PROGRAM Counters
  VAR
    h01_a : BOOL;
    CTU0 : CTU;
    h01_q : BOOL;
    h01_b : BOOL;
    h01_c : BOOL;
    h01_d : BOOL;
    h01_cv : INT;
    h02_a : BOOL;
    CTUD0 : CTUD;
    h02_qu : BOOL;
    h02_b : BOOL;
    h02_c : BOOL;
    h02_d : BOOL;
    h02_e : BOOL;
    h02_g : BOOL;
    h02_f : BOOL;
    h02_h : BOOL;
    h02_i : BOOL;
    h02_k : BOOL;
    h02_j : BOOL;
    h02_qd : BOOL;
    h02_cv : INT;
    h03_a : BOOL;
    SR0 : SR;
    h03_q1 : BOOL;
    h03_c : BOOL;
    h03_b : BOOL;
    h03_d : BOOL;
    h03_e : BOOL;
    RS0 : RS;
    h03_q2 : BOOL;
    h03_f : BOOL;
    h03_h : BOOL;
    h03_g : BOOL;
    h04_e : BOOL;
    TON0 : TON;
    h04_q : BOOL;
    h04_a : BOOL;
    h04_b : BOOL;
    h04_c : BOOL;
    h04_d : BOOL;
    h04_et : TIME;
  END_VAR

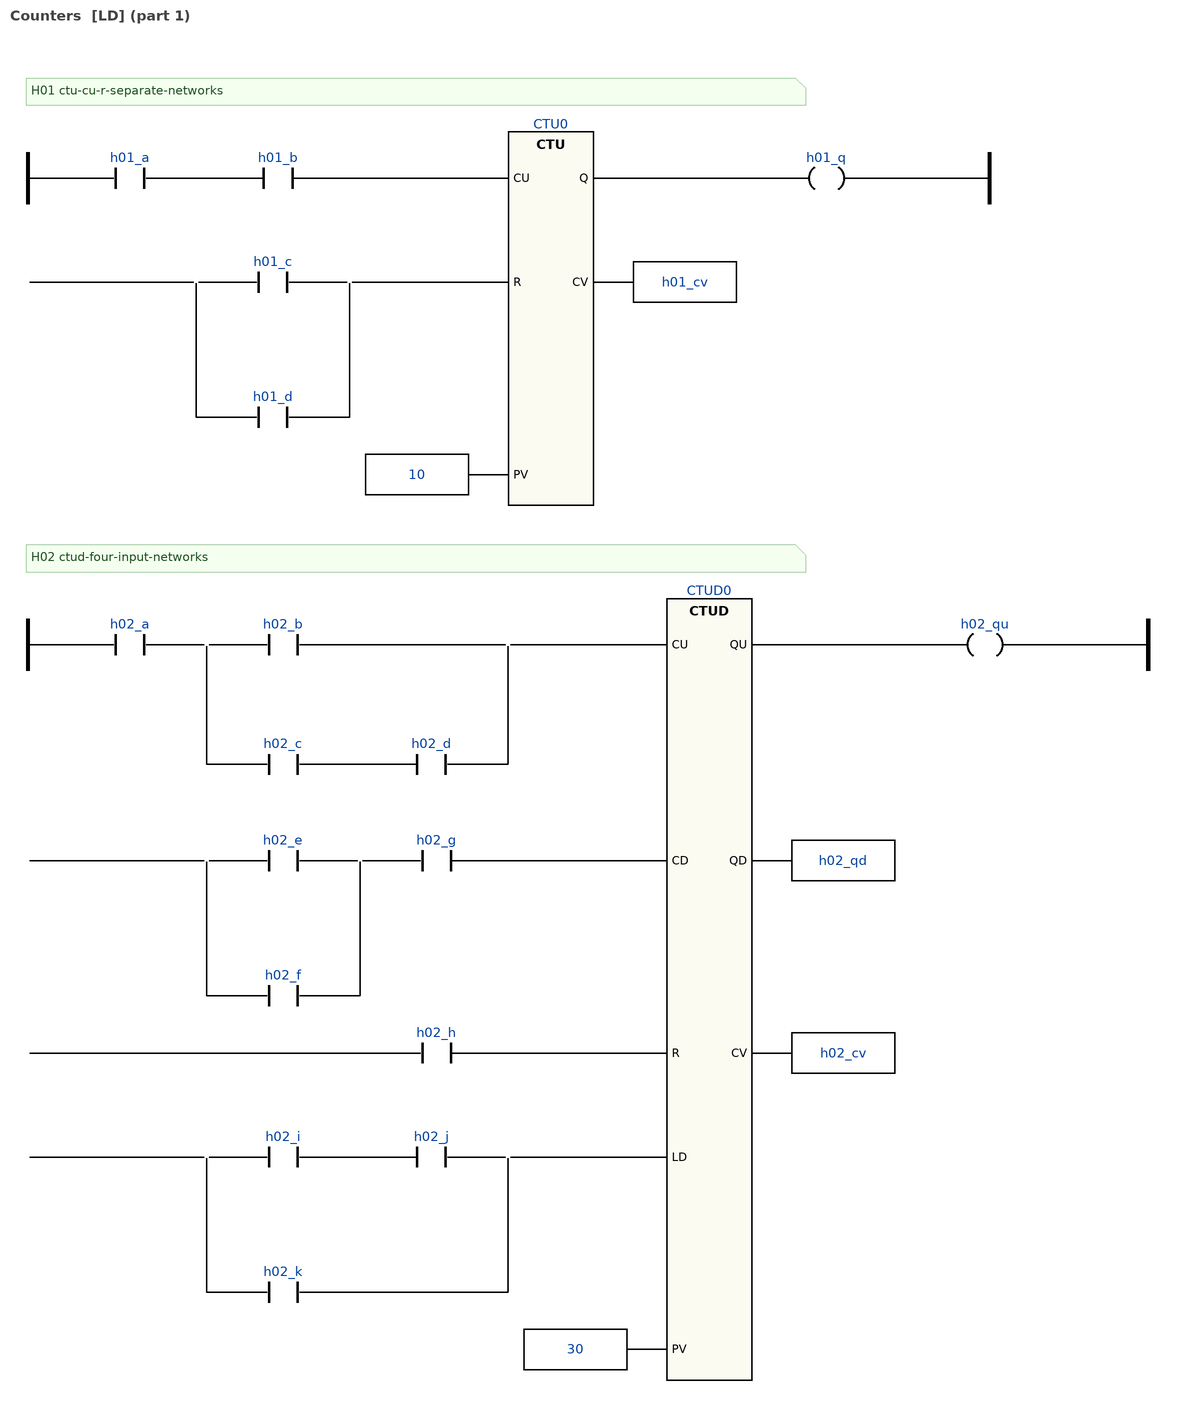
(* LD diagram, written out as Structured Text *)
(* H01 ctu-cu-r-separate-networks *)
CTU0(CU := h01_a AND h01_b, R := h01_c OR h01_d, PV := 10);
h01_q := CTU0.Q;
h01_cv := CTU0.CV;
(* H02 ctud-four-input-networks *)
CTUD0(CU := h02_a AND (h02_b OR h02_c AND h02_d), CD := (h02_e OR h02_f) AND h02_g, R := h02_h, LD := h02_k OR h02_i AND h02_j, PV := 30);
h02_qu := CTUD0.QU;
h02_qd := CTUD0.QD;
h02_cv := CTUD0.CV;
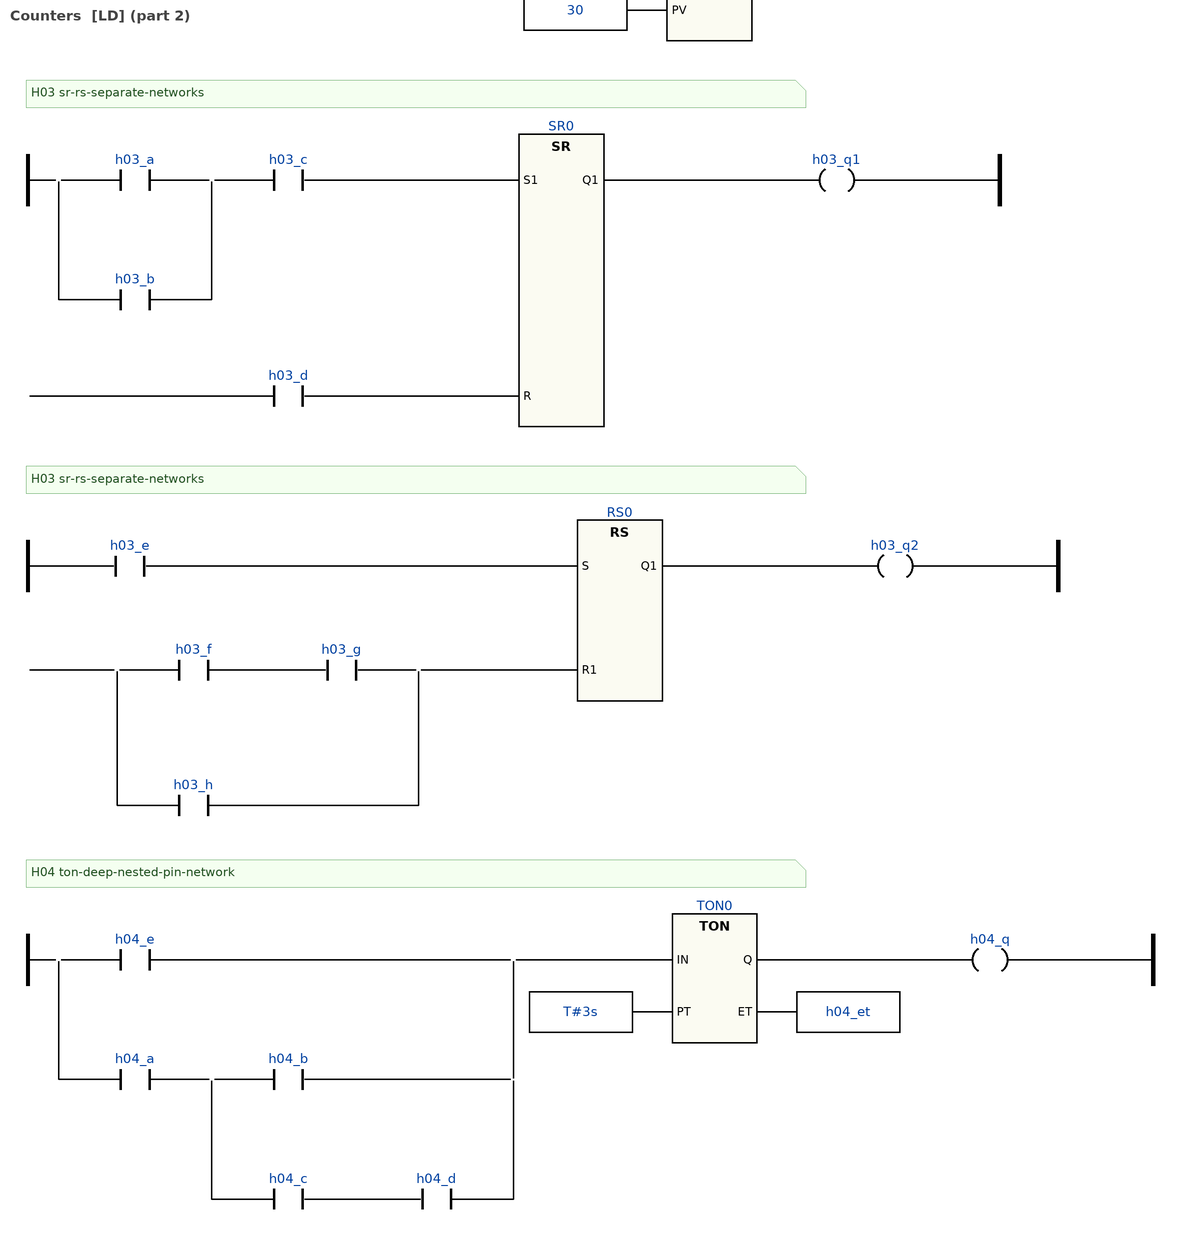
(* H03 sr-rs-separate-networks *)
SR0(S1 := (h03_a OR h03_b) AND h03_c, R := h03_d);
h03_q1 := SR0.Q1;
(* H03 sr-rs-separate-networks *)
RS0(S := h03_e, R1 := h03_h OR h03_f AND h03_g);
h03_q2 := RS0.Q1;
(* H04 ton-deep-nested-pin-network *)
TON0(IN := h04_e OR h04_a AND h04_b OR h04_a AND h04_c AND h04_d, PT := T#3s);
h04_q := TON0.Q;
h04_et := TON0.ET;
END_PROGRAM
